(* PLC project Motor_Control, PLCAutoPilot Machine Expert Logic Builder V19.2.3.0, author PLCAutoPilot *)
(* stored: creationDateTime 2025-12-30T02:10:00.0000000, version 1.0.0.0, modificationDateTime 2025-12-30T02:10:00.0000000 *)

PROGRAM Motor_Control_LD
  VAR
    StartPB AT %IX0.0 : BOOL;
    StopPB AT %IX0.1 : BOOL;
    OverloadTrip AT %IX0.2 : BOOL;
    EmergencyStop AT %IX0.3 : BOOL;
    MotorContactor AT %QX0.0 : BOOL;
    RunIndicator AT %QX0.1 : BOOL;
    FaultIndicator AT %QX0.2 : BOOL;
  END_VAR
  VAR
    MotorRunning : BOOL;
    MotorFault : BOOL;
    SafetyOK : BOOL;
    StartCondition : BOOL;
    StartupTimer : TON;
  END_VAR

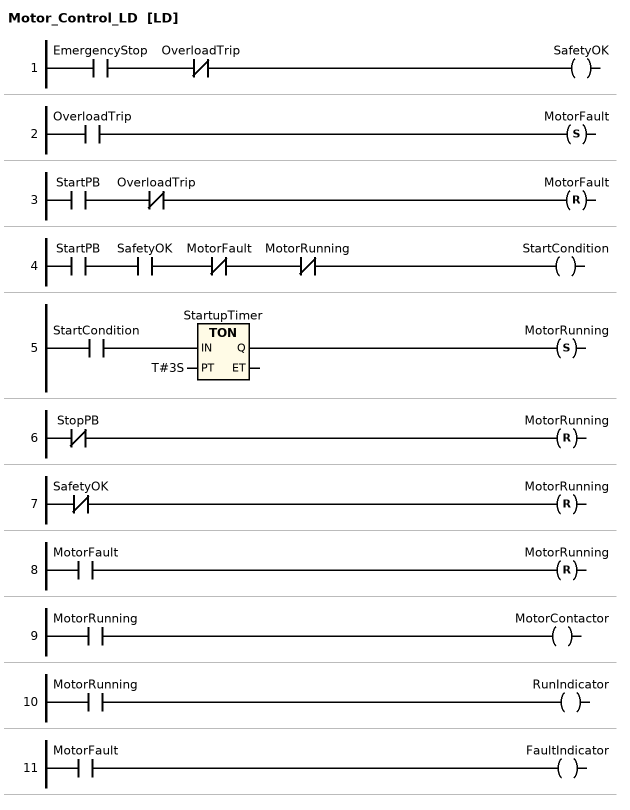
(* LD diagram, written out as Structured Text *)
(* Network 1: Safety Interlock Check *)

SafetyOK := EmergencyStop AND NOT OverloadTrip;
(* Network 2: Fault SET on Overload Trip *)

IF OverloadTrip THEN MotorFault := TRUE; END_IF;
(* Network 3: Fault RESET when Start AND Overload Clear *)

IF StartPB AND NOT OverloadTrip THEN MotorFault := FALSE; END_IF;
(* Network 4: Start Condition = Start AND Safe AND NOT Fault AND NOT Running *)

StartCondition := StartPB AND SafetyOK AND NOT MotorFault AND NOT MotorRunning;
(* Network 5: 3 Second Startup Timer *)

StartupTimer(IN := StartCondition, PT := T#3S);
IF StartupTimer.Q THEN MotorRunning := TRUE; END_IF;
(* Network 6: Motor RESET on Stop Press or Safety Fail *)

IF NOT StopPB THEN MotorRunning := FALSE; END_IF;
(* Network 7: Motor RESET on Safety NOT OK *)

IF NOT SafetyOK THEN MotorRunning := FALSE; END_IF;
(* Network 8: Motor RESET on Fault *)

IF MotorFault THEN MotorRunning := FALSE; END_IF;
(* Network 9: Motor Contactor Output *)

MotorContactor := MotorRunning;
(* Network 10: Run Indicator Lamp *)

RunIndicator := MotorRunning;
(* Network 11: Fault Indicator Lamp *)

FaultIndicator := MotorFault;
END_PROGRAM
